(* IEC 61131-3 sources: codesys-to-s7/tests/corpus/C2S7-POU-FBINFC/pos, 1 file *)

(* ---- input.st ---- *)
FUNCTION F_Case : INT
VAR
    t : TON;
END_VAR
t(IN := TRUE, PT := T#1S); F_Case := 0;
END_FUNCTION
